// 	                                     Level := 4,
// 	                                     Light_Guard_IO:=LIGHT_GUARDS_C2201___CH1,
// 	                                     Light_Guard_Bypass=>Light_Guard_Bypass_2_,
// 	                                     System_Busy:=System_2_Busy);
// 	                110502:
// 	                    Feed_BCNV_Cnv2_1_( System_No := 2,
// 	                                     Level := 5,
// 	                                     Light_Guard_IO:=LIGHT_GUARDS_C2201___CH1,
// 	                                     Light_Guard_Bypass=>Light_Guard_Bypass_2_,
// 	                                     System_Busy:=System_2_Busy);
// 	                110602:
// 	                    Feed_BCNV_Cnv2_1_( System_No := 2,
// 	                                     Level := 6,
// 	                                     Light_Guard_IO:=LIGHT_GUARDS_C2201___CH1,
// 	                                     Light_Guard_Bypass=>Light_Guard_Bypass_2_,
// 	                                     System_Busy:=System_2_Busy);
// 	                110702:
// 	                    Feed_BCNV_Cnv2_1_( System_No := 2,
// 	                                     Level := 7,
// 	                                     Light_Guard_IO:=LIGHT_GUARDS_C2201___CH1,
// 	                                     Light_Guard_Bypass=>Light_Guard_Bypass_2_,
// 	                                     System_Busy:=System_2_Busy);
// 	                110802:
// 	                    Feed_BCNV_Cnv2_1_( System_No := 2,
// 	                                     Level := 8,
// 	                                     Light_Guard_IO:=LIGHT_GUARDS_C2201___CH1,
// 	                                     Light_Guard_Bypass=>Light_Guard_Bypass_2_,
// 	                                     System_Busy:=System_2_Busy);
// 
// 
// 	                100103:
// 	                    Feed_BCNV_Cnv1_1_( System_No := 3,
// 	                                     Level := 1,
// 	                                     Light_Guard_IO:=LIGHT_GUARDS_C3101___CH1,
// 	                                     Light_Guard_Bypass=>Light_Guard_Bypass_3_,
// 	                                     System_Busy:=System_3_Busy);
// 	                100203:
// 	                    Feed_BCNV_Cnv1_1_( System_No := 3,
// 	                                     Level := 2,
// 	                                     Light_Guard_IO:=LIGHT_GUARDS_C3101___CH1,
// 	                                     Light_Guard_Bypass=>Light_Guard_Bypass_3_,
// 	                                     System_Busy:=System_3_Busy);
// 	                100303:
// 	                    Feed_BCNV_Cnv1_1_( System_No := 3,
// 	                                     Level := 3,
// 	                                     Light_Guard_IO:=LIGHT_GUARDS_C3101___CH1,
// 	                                     Light_Guard_Bypass=>Light_Guard_Bypass_3_,
// 	                                     System_Busy:=System_3_Busy);
// 	                100403:
// 	                    Feed_BCNV_Cnv1_1_( System_No := 3,
// 	                                     Level := 4,
// 	                                     Light_Guard_IO:=LIGHT_GUARDS_C3101___CH1,
// 	                                     Light_Guard_Bypass=>Light_Guard_Bypass_3_,
// 	                                     System_Busy:=System_3_Busy);
// 	                100503:
// 	                    Feed_BCNV_Cnv1_1_( System_No := 3,
// 	                                     Level := 5,
// 	                                     Light_Guard_IO:=LIGHT_GUARDS_C3101___CH1,
// 	                                     Light_Guard_Bypass=>Light_Guard_Bypass_3_,
// 	                                     System_Busy:=System_3_Busy);
// 	                100603:
// 	                    Feed_BCNV_Cnv1_1_( System_No := 3,
// 	                                     Level := 6,
// 	                                     Light_Guard_IO:=LIGHT_GUARDS_C3101___CH1,
// 	                                     Light_Guard_Bypass=>Light_Guard_Bypass_3_,
// 	                                     System_Busy:=System_3_Busy);
// 	                100703:
// 	                    Feed_BCNV_Cnv1_1_( System_No := 3,
// 	                                     Level := 7,
// 	                                     Light_Guard_IO:=LIGHT_GUARDS_C3101___CH1,
// 	                                     Light_Guard_Bypass=>Light_Guard_Bypass_3_,
// 	                                     System_Busy:=System_3_Busy);
// 	                100803:
// 	                    Feed_BCNV_Cnv1_1_( System_No := 3,
// 	                                     Level := 8,
// 	                                     Light_Guard_IO:=LIGHT_GUARDS_C3101___CH1,
// 	                                     Light_Guard_Bypass=>Light_Guard_Bypass_3_,
// 	                                     System_Busy:=System_3_Busy);
// 
// 	                110103:
// 	                    Feed_BCNV_Cnv2_1_( System_No := 3,
// 	                                     Level := 1,
// 	                                     Light_Guard_IO:=LIGHT_GUARDS_C3201___CH1,
// 	                                     Light_Guard_Bypass=>Light_Guard_Bypass_3_,
// 	                                     System_Busy:=System_3_Busy);
// 	                110203:
// 	                    Feed_BCNV_Cnv2_1_( System_No := 3,
// 	                                     Level := 2,
// 	                                     Light_Guard_IO:=LIGHT_GUARDS_C3201___CH1,
// 	                                     Light_Guard_Bypass=>Light_Guard_Bypass_3_,
// 	                                     System_Busy:=System_3_Busy);
// 	                110303:
// 	                    Feed_BCNV_Cnv2_1_( System_No := 3,
// 	                                     Level := 3,
// 	                                     Light_Guard_IO:=LIGHT_GUARDS_C3201___CH1,
// 	                                     Light_Guard_Bypass=>Light_Guard_Bypass_3_,
// 	                                     System_Busy:=System_3_Busy);
// 	                110403:
// 	                    Feed_BCNV_Cnv2_1_( System_No := 3,
// 	                                     Level := 4,
// 	                                     Light_Guard_IO:=LIGHT_GUARDS_C3201___CH1,
// 	                                     Light_Guard_Bypass=>Light_Guard_Bypass_3_,
// 	                                     System_Busy:=System_3_Busy);
// 	                110503:
// 	                    Feed_BCNV_Cnv2_1_( System_No := 3,
// 	                                     Level := 5,
// 	                                     Light_Guard_IO:=LIGHT_GUARDS_C3201___CH1,
// 	                                     Light_Guard_Bypass=>Light_Guard_Bypass_3_,
// 	                                     System_Busy:=System_3_Busy);
// 	                110603:
// 	                    Feed_BCNV_Cnv2_1_( System_No := 3,
// 	                                     Level := 6,
// 	                                     Light_Guard_IO:=LIGHT_GUARDS_C3201___CH1,
// 	                                     Light_Guard_Bypass=>Light_Guard_Bypass_3_,
// 	                                     System_Busy:=System_3_Busy);
// 	                110703:
// 	                    Feed_BCNV_Cnv2_1_( System_No := 3,
// 	                                     Level := 7,
// 	                                     Light_Guard_IO:=LIGHT_GUARDS_C3201___CH1,
// 	                                     Light_Guard_Bypass=>Light_Guard_Bypass_3_,
// 	                                     System_Busy:=System_3_Busy);
// 	                110803:
// 	                    Feed_BCNV_Cnv2_1_( System_No := 3,
// 	                                     Level := 8,
// 	                                     Light_Guard_IO:=LIGHT_GUARDS_C3201___CH1,
// 	                                     Light_Guard_Bypass=>Light_Guard_Bypass_3_,
// 	                                     System_Busy:=System_3_Busy);
// 
// 
// 	                100104:
// 	                    Feed_BCNV_Cnv1_1_( System_No := 4,
// 	                                     Level := 1,
// 	                                     Light_Guard_IO:=TRUE,
// 	                                     Light_Guard_Bypass=>No_Light_Guard,
// 	                                     System_Busy:=System_4_Busy);
// 	                100204:
// 	                    Feed_BCNV_Cnv1_1_( System_No := 4,
// 	                                     Level := 2,
// 	                                     Light_Guard_IO:=TRUE,
// 	                                     Light_Guard_Bypass=>No_Light_Guard,
// 	                                     System_Busy:=System_4_Busy);
// 	                100304:
// 	                    Feed_BCNV_Cnv1_1_( System_No := 4,
// 	                                     Level := 3,
// 	                                     Light_Guard_IO:=TRUE,
// 	                                     Light_Guard_Bypass=>No_Light_Guard,
// 	                                     System_Busy:=System_4_Busy);
// 	                100404:
// 	                    Feed_BCNV_Cnv1_1_( System_No := 4,
// 	                                     Level := 4,
// 	                                     Light_Guard_IO:=TRUE,
// 	                                     Light_Guard_Bypass=>No_Light_Guard,
// 	                                     System_Busy:=System_4_Busy);
// 	                100504:
// 	                    Feed_BCNV_Cnv1_1_( System_No := 4,
// 	                                     Level := 5,
// 	                                     Light_Guard_IO:=TRUE,
// 	                                     Light_Guard_Bypass=>No_Light_Guard,
// 	                                     System_Busy:=System_4_Busy);
// 	                100604:
// 	                    Feed_BCNV_Cnv1_1_( System_No := 4,
// 	                                     Level := 6,
// 	                                     Light_Guard_IO:=TRUE,
// 	                                     Light_Guard_Bypass=>No_Light_Guard,
// 	                                     System_Busy:=System_4_Busy);
// 	                100704:
// 	                    Feed_BCNV_Cnv1_1_( System_No := 4,
// 	                                     Level := 7,
// 	                                     Light_Guard_IO:=TRUE,
// 	                                     Light_Guard_Bypass=>No_Light_Guard,
// 	                                     System_Busy:=System_4_Busy);
// 	                100804:
// 	                    Feed_BCNV_Cnv1_1_( System_No := 4,
// 	                                     Level := 8,
// 	                                     Light_Guard_IO:=TRUE,
// 	                                     Light_Guard_Bypass=>No_Light_Guard,
// 	                                     System_Busy:=System_4_Busy);
// 
// 	                120005:
// 	                    Feed_ECNV_1_( System_No := 5);
// 
// 	                100105:
// 	                    Feed_BCNV_Cnv1_1_( System_No := 5,
// 	                                     Level := 1,
// 	                                     Light_Guard_IO:=TRUE,
// 	                                     Light_Guard_Bypass=>No_Light_Guard,
// 	                                     System_Busy:=System_5_Busy);
// 	                100205:
// 	                    Feed_BCNV_Cnv1_1_( System_No := 5,
// 	                                     Level := 2,
// 	                                     Light_Guard_IO:=TRUE,
// 	                                     Light_Guard_Bypass=>No_Light_Guard,
// 	                                     System_Busy:=System_5_Busy);
// 	                100305:
// 	                    Feed_BCNV_Cnv1_1_( System_No := 5,
// 	                                     Level := 3,
// 	                                     Light_Guard_IO:=TRUE,
// 	                                     Light_Guard_Bypass=>No_Light_Guard,
// 	                                     System_Busy:=System_5_Busy);
// 	                100405:
// 	                    Feed_BCNV_Cnv1_1_( System_No := 5,
// 	                                     Level := 4,
// 	                                     Light_Guard_IO:=TRUE,
// 	                                     Light_Guard_Bypass=>No_Light_Guard,
// 	                                     System_Busy:=System_5_Busy);
// 	                100505:
// 	                    Feed_BCNV_Cnv1_1_( System_No := 5,
// 	                                     Level := 5,
// 	                                     Light_Guard_IO:=TRUE,
// 	                                     Light_Guard_Bypass=>No_Light_Guard,
// 	                                     System_Busy:=System_5_Busy);
// 	                100605:
// 	                    Feed_BCNV_Cnv1_1_( System_No := 5,
// 	                                     Level := 6,
// 	                                     Light_Guard_IO:=TRUE,
// 	                                     Light_Guard_Bypass=>No_Light_Guard,
// 	                                     System_Busy:=System_5_Busy);
// 	                100705:
// 	                    Feed_BCNV_Cnv1_1_( System_No := 5,
// 	                                     Level := 7,
// 	                                     Light_Guard_IO:=TRUE,
// 	                                     Light_Guard_Bypass=>No_Light_Guard,
// 	                                     System_Busy:=System_5_Busy);
// 	                100805:
// 	                    Feed_BCNV_Cnv1_1_( System_No := 5,
// 	                                     Level := 8,
// 	                                     Light_Guard_IO:=TRUE,
// 	                                     Light_Guard_Bypass=>No_Light_Guard,
// 	                                     System_Busy:=System_5_Busy);
// 	            END_CASE;
// 	        END_IF;
// 
// 
// 	T_Reset_Charge.TON(IN := Screen_DB.Charge_VTD OR Screen_DB.Charge_Cnv OR Screen_DB.Charge_VTD_Commands OR Screen_DB.Charge_Cnv_Commands,
// 	                       PT := T#2S);
// 
// 	   IF T_Reset_Charge.Q THEN
// 	    Screen_DB.Charge_VTD := FALSE;
// 	    Screen_DB.Charge_Cnv := FALSE;
// 	    Screen_DB.Charge_VTD_Commands := FALSE;
// 	    Screen_DB.Charge_Cnv_Commands := FALSE;
// 	END_IF;

END_FUNCTION_BLOCK

(* stored: Version 1.1.0.1
   POU Conveyor_HMI_FB: Id {f566d77c-2b55-5962-b9fe-d6593304177f}, SpecialFunc None *)
